(* IEC 61131-3 sources: iFA_git_test/GIT test/PLC_2/Programs, 2 files *)

(* ---- DefaultVariableTable.st ---- *)
(*NodeCRC64:15794442468608431415, FileCRC64:15794442468608431415*)
VAR_GLOBAL
END_VAR
(*{"Version":"1.0.0.0","Path":"Default_variable_table","ObjectType":"Global"}*)
END_VAR_GLOBAL

(* ---- Main.st ---- *)
(*NodeCRC64:4207710498223751431, FileCRC64:4207710498223751431*)
PROGRAM Main
VAR
END_VAR
Body

EndBody
(*{"Version":"1.0.0.0","Path":"Main","ObjectType":"Program"}*)
END_PROGRAM
